TYPE ST_Polynom5Factor :
STRUCT
	fA0: LREAL;
	fA1: LREAL;
	fA2: LREAL;
	fA3: LREAL;
	fA4: LREAL;
	fA5: LREAL;
END_STRUCT
END_TYPE

(* stored: Version 1.1.0.1, ProductVersion 3.1.4024.12
   DUT ST_Polynom5Factor: Id {88261255-1c8e-4d92-b737-7495bd943038} *)
